Fanuc KAREL source: kb00048.KL

-- PROVISIONAL review KL for V1013-1; original PC SHA256 24a985340a15fb620e574c03ec45e26baf0dbaac37921a871b4703c9454e37da
-- Incomplete behavior may be omitted. Consult companion uncertainty JSON. Do not deploy.
PROGRAM KB00048
%NOLOCKGROUP
VAR
  P1 : REAL
  RESULT : REAL
BEGIN
  -- UNRESOLVED_PC offsets 5-16; opcodes 2E,23
  -- UNRESOLVED_PC offsets 21-36; opcodes 27,22,76,23
  -- UNRESOLVED_PC offsets 41-45; opcodes 7F
END KB00048
